Yaskawa INFORM job: LONGPRO4.JBI

/JOB
//NAME LONGPRO4
//POS
///NPOS 5,0,0,0,0,0
///TOOL 9
///POSTYPE PULSE
///PULSE
C00000=0,-10240,0,-34475,0,0,22983
C00001=20480,-10240,0,-34475,0,-8704,22983
C00002=0,-10240,0,-34475,0,0,22983
C00003=20480,-10240,0,-34475,0,-8704,22983
C00004=0,-10240,0,-34475,0,0,22983
//INST
<volatile>
///COMM Generated using RoboDK
///ATTR SC,RW
///GROUP1 RB1
NOP
MOVJ C00000 VJ=50.00
MOVJ C00001 VJ=50.00
MOVJ C00002 VJ=50.00
MOVJ C00003 VJ=50.00
MOVJ C00004 VJ=50.00
END
